(* IEC 61131-3 sources: 89152_FlorisHendrix_AfstudeerProject/89152_FlorisHendrix_ExamenProject/Stations/MachineControl/MachineControl/Network/HW_Network, 1 file *)

(* ---- ONE_HW_Network_Table.st ---- *)
#define OBJECTS_CONFIG

//Define part of class SdiasBase
//Address to access the Dataobject list via SPI SDO Read
#define SDIAS_SPI_DATA_OBJECT_LIST_PAGE_ADDRESS               16#FFFF
#define SDIAS_SPI_DATA_OBJECT_LIST_PAGE_OFFSET                16#00
#define SDIAS_SPI_DATA_OBJECT_LIST_IDENTIFIER                 16#12345678

//Defines the number of optional list elements in the SPI List

#define SDIAS_SPI_NUMBER_OF_OPTIONAL_ELEMENTS                 16

#define SDIAS_SPI_HEADER_BEFORE_OPTIONAL_ELEMENTS             16#18
#define SDIAS_SPI_HARDWARE_VERSION_OFFSET                     16#C
#define SDIAS_SPI_VENDOR_ID_OFFSET                            16#0

#define SDIAS_SPI_MASTER_ADRESS_TRANSMIT_BUFFER0              16#0000
#define SDIAS_SPI_MASTER_ADRESS_TRANSMIT_BUFFER1              16#0080
#define SDIAS_SPI_MASTER_ADRESS_RECEIVE_BUFFER0               16#0000
#define SDIAS_SPI_MASTER_ADRESS_RECEIVE_BUFFER1               16#0080
#define SDIAS_SPI_MASTER_ADRESS_PAGE_ADRESS                   16#0100
#define SDIAS_SPI_MASTER_ADRESS_PREDEFINED_COMMAND_REGISTER   16#0102
#define SDIAS_SPI_MASTER_ADRESS_SINGLE_COMMAND_REGISTER       16#0103
#define SDIAS_SPI_MASTER_ADRESS_STATUS_REGISTER               16#0104
#define SDIAS_SPI_MASTER_ADRESS_REQUEST_REGISTER              16#0105
#define SDIAS_SPI_MASTER_ADRESS_GRANT_REGISTER                16#0106
#define SDIAS_SPI_MASTER_ADRESS_CLEAR_REQUEST_REGISTER        16#0107
#define SDIAS_SPI_MASTER_ADRESS_FEATURE_REGISTER              16#0108

#define SDIAS_SPI_MASTER_SOFTWARE_REQUEST                     1

#define SDIAS_SPI_MASTER_COMMAND_PAGE_READ                    16#01
#define SDIAS_SPI_MASTER_COMMAND_PAGE_PROGRAM                 16#02
#define SDIAS_SPI_MASTER_COMMAND_SECTOR_ERASE                 16#03
#define SDIAS_SPI_MASTER_COMMAND_REBOOT_FPGA                  16#F0

#define SDIAS_SPI_MASTER_STATE_BUSY                           16#00
#define SDIAS_SPI_MASTER_STATE_READY                          16#01

#define SDIAS_SPI_SECTOR_SIZE                                 65536 // 256*256
#define SDIAS_SPI_PAGE_SIZE                                   256

#define SDIAS_SPI_WRITE_MAX_RETRIES                           2
#define SDIAS_SPI_TIMEOUT                                     500  //timeout for spi accesses
#define SDIAS_SPI_LOCK_TIMEOUT                                6   //this value is multiplied with the buscycletime [µs] (6*1000=6.000 msec timeout)

//SPI List IDs
#define SDIAS_SPI_IDENTIFICATION_LIST_ID  1
#define SDIAS_SPI_FLASH_CONFIGURATION_ID  2
#define SDIAS_SPI_VENDOR_NAME_ID          3
#define SDIAS_SPI_DEVICE_NAME_ID          4
#define SDIAS_SPI_SERIAL_NUMBER_ID        5
#define SDIAS_SPI_ORDERING_NUMBER_ID      6
#define SDIAS_SPI_DOCUMENTATION_PDF_ID    7
#define SDIAS_SPI_CALIB_DATA_ID           10
#define SDIAS_SPI_PDO_INFORMATION_ID      128

//SPI Access
#define SDIAS_SPI_ACCESS_ID_HW_TREE          1
#define SDIAS_SPI_ACCESS_ID_HWK_INTERNAL     2
#include "..\..\Class\SdiasManager\SdiasManager.h"
#include "..\..\Class\SdiasBase\SdiasBase.h"
#include "..\..\Class\HwControl\HwControl.h"
#include "..\..\Source\interfaces\lsl_st_hardwaretree.h"
#include "..\..\Source\interfaces\lsl_st_mt.h"
//Define part of class _BusInterfaceSdiasDriveMng
#define BUSIF_SDIASDRIVEMNG_OFFSET_TYPELABEL        0x0000
#define BUSIF_SDIASDRIVEMNG_PARALIST_INDEX_SET      0x2210
#define BUSIF_SDIASDRIVEMNG_PARALIST_INDEX_INFO     0x2211
#define BUSIF_SDIASDRIVEMNG_PARALIST_INDEX_SETNR    174

#define BUSIF_SDIASDRIVEMNG_MAX_SERVICEBOX          4
#define BUSIF_SDIASDRIVEMNG_SDO_RESPONSE_TIMEOUT    SDIAS_SDO_TIMEOUT * 2
#define BUSIF_SDIASDRIVEMNG_SDO_TYPELABEL_TIMEOUT   10000  //10 sec timeout to read typelabel

#define BUSIF_SDIASDRIVEMNG_SDO_SERVICE_APP_MDD100        0x4150
#define BUSIF_SDIASDRIVEMNG_SDO_SERVICE_APP_LASAL         0x4C41
#define BUSIF_SDIASDRIVEMNG_SDO_SERVICE_APP_CANOPEN       0x4453
#define BUSIF_SDIASDRIVEMNG_SDO_SERVICE_APP_CANOPEN_LASAL 0x444C

#define BUSIF_SDIASDRIVEMNG_FULL_PARADATA_SIZE   12
#define BUSIF_SDIASDRIVEMNG_CANOPEN_FOOTER_SIZE   4
#define BUSIF_SDIASDRIVEMNG_LASAL_PARADATA_SIZE   4

// if it's an sr011 or sr012 module we must set the pll system periode time with this offset
#define BUSIF_SDIASDRIVEMNG_SR01X_PLL_OFFSET    16#140
#include "..\..\class\_drivemngbase\drivemngbase.h"
//Define part of class _DriveAxisBase
// Device ID for the Drive Cards
#define DRIVEMNG_AXISDEVICEID_SDD_OFFSET         0
#define DRIVEMNG_AXISEVICEID_MDD_OFFSET   16#10000
#define DRIVEMNG_AXISEVICEID_SDIAS_OFFSET 16#20000

#define DRIVEAXIS_SPEED_SFFLIMITATION_USERINFO_0   32767
#define DRIVEAXIS_SPEED_SFFLIMITATION_USERINFO_1    1000
#define DRIVEAXIS_TORQUE_LIMITATION_VALUE           1000
#include "..\..\Class\_DriveMngBase\SDDDefinitions.h"
#include "..\..\Class\_DriveAxisBase\_DriveAxis_A_INT_Def.h"
//Define part of class _DriveMngBase
#ifndef _T_DRIVEMNGBASE_H
#define _T_DRIVEMNGBASE_H

// DiasDrive Constants
#DEFINE SDDMAXENTRIES   32        // maximale Anzahl an Achsen
#DEFINE SDDMAXPLACE     3         // maximale Anzahl an Achsen pro Steckplatz

// Device ID for the Drive IF Cards
#define DRIVEMNG_BUSDEVICEID_VAC011    11
#define DRIVEMNG_BUSDEVICEID_VAC012  1061
#define DRIVEMNG_BUSDEVICEID_VAC013  1075

#define DRIVEMNG_BUSDEVICEID_MDD     1071

// Device ID for the Drive Cards
#define DRIVEMNG_DRVDEVICEID_SDD_OFFSET 0

#define DRIVEMNG_DRVDEVICEID_SDD305 DRIVEMNG_DRVDEVICEID_SDD_OFFSET + 16
#define DRIVEMNG_DRVDEVICEID_SDD310 DRIVEMNG_DRVDEVICEID_SDD_OFFSET +  3
#define DRIVEMNG_DRVDEVICEID_SDD315 DRIVEMNG_DRVDEVICEID_SDD_OFFSET +  1
#define DRIVEMNG_DRVDEVICEID_SDD335 DRIVEMNG_DRVDEVICEID_SDD_OFFSET + 12

#define DRIVEMNG_DRVDEVICEID_SDD205 DRIVEMNG_DRVDEVICEID_SDD_OFFSET + 22
#define DRIVEMNG_DRVDEVICEID_SDD210 DRIVEMNG_DRVDEVICEID_SDD_OFFSET +  9
#define DRIVEMNG_DRVDEVICEID_SDD215 DRIVEMNG_DRVDEVICEID_SDD_OFFSET +  5

#define DRIVEMNG_DRVDEVICEID_SDD105 DRIVEMNG_DRVDEVICEID_SDD_OFFSET + 21
#define DRIVEMNG_DRVDEVICEID_SDD115 DRIVEMNG_DRVDEVICEID_SDD_OFFSET + 10
#define DRIVEMNG_DRVDEVICEID_SDD120 DRIVEMNG_DRVDEVICEID_SDD_OFFSET +  7

#define DRIVEMNG_DRVDEVICEID_MDD_OFFSET 16#10000

#define DRIVEMNG_DRVDEVICEID_MDD111 DRIVEMNG_DRVDEVICEID_MDD_OFFSET + 1
#define DRIVEMNG_DRVDEVICEID_MDD121 DRIVEMNG_DRVDEVICEID_MDD_OFFSET + 2

#define DRIVEMNG_DRVDEVICEID_SDIAS_OFFSET 16#20000

#define DRIVEMNG_DRVDEVICEID_DC061 DRIVEMNG_DRVDEVICEID_SDIAS_OFFSET + 16#180 // 1 = 1 Achse 80 SDIAS

#define DRIVEMNG_DRIVESCOPE_GETALL_PARAM    16#2080
#define DRIVEMNG_DRIVESCOPE_SCOPE_BIT       16#60000000
#define DRIVEMNG_DRIVESCOPE_SINDEX_RANGE    511

#define DRIVEMNG_DEFAULT_CPU_LOGFILENAME_PATH           "C:\sysmsg\DriveLog"
#define DRIVEMNG_DEFAULT_CPU_DEBUGLOGFILENAME_PATH      "C:\sysmsg\DriveDebugLog"
#define DRIVEMNG_DEFAULT_CPU_LOGFILENAME_EXTENSION      ".txt"

#define DRIVEMNG_DEFAULT_DRIVE_LOGFILENAME_PATH         "C:\"
#define DRIVEMNG_DEFAULT_DRIVE_LOGFILENAME_NAME         "DriveLog.txt"
#define DRIVEMNG_DEFAULT_DRIVE_DEBUGLOGFILENAME_NAME    "DriveDebugLog.txt"

#define DRIVEMNG_FILE_HANDLING_RETCODE_NOERROR                    0
#define DRIVEMNG_FILE_HANDLING_RETCODE_FILEHANDLING_BUSY         -2   // = DRIVEVVBASE_VANDAL_FILEHANDLING_ERROR_BUSY -2
#define DRIVEMNG_FILE_HANDLING_RETCODE_CMDVERSION_NOTSUPPORTED  -92
#define DRIVEMNG_FILE_HANDLING_RETCODE_WRITEPARA_FAILED         -93
#define DRIVEMNG_FILE_HANDLING_RETCODE_WRITEPARA_TIMEOUT        -94
#define DRIVEMNG_FILE_HANDLING_RETCODE_READBACKPARA_FAILED      -95
#define DRIVEMNG_FILE_HANDLING_RETCODE_READBACKPARA_TIMEOUT     -96
#define DRIVEMNG_FILE_HANDLING_RETCODE_AXIS_ENABLED             -97
#define DRIVEMNG_FILE_HANDLING_RETCODE_NOT_ONLINE               -98
#define DRIVEMNG_FILE_HANDLING_RETCODE_NOT_SUPPORTED            -99

#define DRIVEMNG_FILE_HANDLING_TIMEOUT_LOG_PARAM          10000

#define DRIVEMNG_FILESELECT_LOGFILE       0
#define DRIVEMNG_FILESELECT_DEBUGLOGFILE  1

#define DRIVEMNG_FILE_RESERVE_IDFREE         0
#define DRIVEMNG_FILE_RESERVE_IDDEFAULT     10
#define DRIVEMNG_FILE_RESERVE_IDGETLOGFILE  20

#endif // _T_DRIVEMNGBASE_H
//Define part of class AI043
#define DEVICE_ID_AI043 1045

#define AI043_ADDR_CYC_WRITE        16#000
#define AI043_ADDR_CYC_READ         16#080
#define AI043_ADDR_CFG_FIRMWARE     16#100
#define AI043_ADDR_STATE_FIRMWARE   16#180

#define AI043_SDO_RESPONSE_TIMEOUT  SDIAS_SDO_TIMEOUT * 2

#define AI043_KTY84_RAW_VALUES_FW_VER_AVAILABLE  16#110
#define AI043_AMOUNT_OF_VALID_CFG   25
#define AI043_AMOUNT_OF_VALID_CFGS_BEFORE_KTY84_ADDED 23

#define AI043_NUMBER_OF_ANALOG_IN   4
#define AI043_INVALID_VALUE         16#80000010$DINT
#define AI043_CABLE_BREAK_MASK      16#0F  //4 BITS

#define AI043_FIRMWARE_MIN          0
#define AI043_FIRMWARE_MAX_CFG12    2500
#define AI043_FIRMWARE_MAX_CFG13    5000
#define AI043_FIRMWARE_MAX_CFG14    10000
#define AI043_FIRMWARE_MAX_CFG15    25000
#define AI043_FIRMWARE_MAX_CFG16    50000
//Define part of class BusInterfaceSDIASInternal
#define BUSIF_INTERNAL_MAX_NR_DO 100

// Defines for Mutex Generation
#define INTERNAL_STR_MUTEX_NAME_SEPERATOR ".."
#define INTERNAL_MUTEX_NAME_END_LENGTH 5
#define INTERNAL_MUTEX_NAME_MAX_LENGTH 32
#include "..\..\Source\BusInterface.h"
//Define part of class Varan_Base
#ifndef _T_VARANBASE_H
#define _T_VARANBASE_H

#define	VARAN_PLL_OFFSET		16#0140
#define VARAN_MULTIPLE_OFFSET	16#01AC

// version of serial number validation (16#10 = 1.0)
#define SERNO_VALIDATION_VERSION 16#10

#define IsTransparent_IS_AVAILABLE

// Defines for Mutex Generation
#define VARAN_STR_MUTEX_NAME_SEPERATOR ".."
#define VARAN_MUTEX_NAME_END_LENGTH 5
#define VARAN_MUTEX_NAME_MAX_LENGTH 32

#define VARAN_SPI_IDENT_LICENCENO_OFFSET    16#14
#define VARAN_SPI_IDENT_HARDWAREVER_OFFSET  16#18

#endif // _T_VARANBASE_H
//Define part of class BusInterfaceVARAN
#define BUSIF_VARAN_MAX_NR_DO     100
#define BUSIF_VARAN_MAX_NR_MOVEDO 100

#define BUSIF_VARAN_MAX_SDO 1

#define BUSIF_VARAN_BUS_READY_VER 16#1109
#include "..\..\Source\interfaces\lsl_st_pci.h"
//Define part of class DM081
#define DEVICE_ID_DM081 1028
//Define part of class DM161
#define DEVICE_ID_DM161 1029
#include "..\..\Class\HwControl\watchdog.h"
#include "..\..\Source\interfaces\lsl_st_sysinfo.h"
#include "..\..\Source\interfaces\lsl_st_systrace.h"
#include "..\..\Class\HwControl\_HWKScope.h"
#include <.\lsl_st_mt.h>
//Define part of class SafetyUDP
#define SAFETY_UDP_MAX_SOCKETS                6     // Max number of socket

#define SAFETY_UDP_CLT_SEND_OK                0    // Send ok
#define SAFETY_UDP_CLT_INVALID_HANDLE        -1    // Invalid handle
#define SAFETY_UDP_CLT_NOT_OPEN              -2    // Socket is not open
#define SAFETY_UDP_CLT_SEND_FAILED           -3    // Send failed
#define SAFETY_UDP_CLT_SEND_BUFFER_FULL      -4    // Send buffer is full
#define SAFETY_UDP_CLT_DATA_TO_BIG           -5    // Data to big

#define SAFETY_UDP_MAXIMUM_SEGMENT_SIZE    1452    // Maximum of user data

#define SAFETY_UDP_TIMEOUT_OPENSOCKET    (1000)    //timeout for opening socket

#define SAFETY_UDP_RECEIVE_TIMEOUT          800

#define SAFETY_UDP_TX_BUFFER_SIZE          1024
//Define part of class SafetyManager
#define LogBufferSize 1000
#include "..\..\Class\SafetyManager\SafetyManager.h"
#include "..\..\Source\interfaces\lsl_st_safetydll.h"
//Define part of class SdiasManager
#define SDIAS_SDO_MAX_LENGTH              128
#define SDIAS_SDO_RINGBUFFER_NO            64
#define SDIAS_SDO_CHANNEL_NO                3   // fixed in the VI hardware to be 3

// watchdog trigger interval (after 130ms of no trigger the SDIAS HW goes into reset again and takes at least another 10ms to be ready again)
#define SDIAS_WATCHDOG_TRIGGER_TIME        40

// time needed by sdias modules to start up after the watchdog is triggered the first time in ms
#define SDIAS_HARDWARE_STARTUP_TIME        15

// sdias manager needs 2 ticks to handle event for read task (measure sync time)
#define SDIAS_SYNC_MEASURE_TICKS            2

// after activating the PLL SyncOut it takes 3 cycles until the SDIAS sync can be injected
#define SDIAS_CYCLES_WAIT_AFTER_SYNC_ENABLE 3

// wait 1 bus cycle at start to get valid numbers in the task info
#define SDIAS_TASKINFO_READY_TICKS          1

// time to wait (in ms) until other tasks in the same or lower priority than post init have done their stuff
#define SDIAS_WAIT_TIME_IN_POST_INIT        1

#define SIZE_PER_SDIAS_CLIENT               16#0400

// for far memory accesses: 1 module can hold maximum 256 1K blocks (0-255)
#define SDIAS_1K_BLOCK_NO                       256

// far memory accesses maximum length in bytes
#define SDIAS_MAX_SIZE_FAR_MEM_ACCESS           127

#define SDIAS_OFFSET_HW_CONFIG              16#FF00
#define SDIAS_OFFSET_TASK_EVENT_IDS         16#FF10
#define SDIAS_OFFSET_FEATURE_INFO           16#FF18
#define SDIAS_OFFSET_APPLI_LED_STATES       16#FF20
#define SDIAS_OFFSET_SYNC_INJECTION_CFG     16#FF3D
#define SDIAS_OFFSET_TRIGGER_UNIT_SETUP_0   16#FF41
#define SDIAS_OFFSET_TRIGGER_UNIT_SETUP_1   16#FF45
#define SDIAS_OFFSET_TASK_START_CFG_0       16#FF60
#define SDIAS_OFFSET_TASK_CONFIG_0          16#FF86
#define SDIAS_OFFSET_TASK_CONFIG_1          16#FF96
#define SDIAS_OFFSET_TASK_INFO_1            16#FF94
#define SDIAS_OFFSET_TASK_HANDSHAKE_1       16#FF9B
#define SDIAS_OFFSET_TASK_DURATION_TIME_1   16#FF9C
#define SDIAS_OFFSET_TASK_DURATION_TIME_2   16#FFAC
#define SDIAS_OFFSET_TASK_CONFIG_2          16#FFA6

#define SDIAS_RETRIES_ALLOWED         2

// mask to get global error flag out of message counter byte of SDO responses
#define SDIAS_MASK_GLOBAL_ERROR_FLAG        16#80

// mask to get message counter out of message counter byte of SDO responses
#define SDIAS_MASK_MESSAGE_COUNTER          16#3F

#define SDIAS_EVENT_MASK_ID_SYNC_OUT0       16#10
#define SDIAS_EVENT_MASK_ID_SYNC_OUT1       16#11
#define SDIAS_EVENT_MASK_ID_SYNC_OUT2       16#12
#define SDIAS_EVENT_MASK_ID_SYNC_OUT3       16#13

#define SDIAS_MANAGER_SYNC_SYNCOUT_ID       16#85
#define SDIAS_TASK_START_EVENT_SYNCOUT_ID   16#86

#define SDIAS_PLACE_NO_MODULE_ADDED_SO_FAR  16#80000000

#define SDIAS_TRIGGER_UNIT_BYTE_SIZE        2

#define SDIAS_WAIT_TIME_FIRMWARE_HANDSHAKE  5 * 1000

// if the firmware version is below this, there might be problems with SCP111 and other modules => print warning at startup
#define SDIAS_FW_VERSION_SDO_ERROR_FIXED    16#120

// if the protocol version ist below this, Control Read/Broadcast Write Command is not supported by sdiasmanager
#define SDIAS_PROTOCOLVERSION_BROADCAST     16#120

// if the cil version ist below this, Control Read/Broadcast Write Command is not supported by OS for local SDIAS.
#define SDIAS_CILVERSION_BROADCAST         16#5001

// timeout for blocking the init during initialisation (in ms)
#define SDIAS_INIT_BLOCK_TIMEOUT            20 * 1000

#define SDIAS_MUTEX_NAME_END_LENGTH 3
#define SDIAS_MUTEX_NAME_MAX_LENGTH 32
#define SDIAS_MUTEX_STR_SEPERATOR   ".."

//#define SDIAS_RT_TIME_MEASUREMENT
#ifdef SDIAS_RT_TIME_MEASUREMENT
  #pragma message("ATTENTION: SDIAS real time measurement is active and needs additional ressources in the realtime task")
#endif

(* SDIAS data object commands  *)
#define	 SDIAS_CMD_END							  0x00			(* End command										          *)
#define	 SDIAS_CMD_ACC_MEMORY				  0x01			(* Access dpram memory								      *)
#define	 SDIAS_CMD_ACC_CONTROL				0x02			(* Access dpram control memory						  *)
#define	 SDIAS_CMD_GLOBAL						  0x03			(* SDIAS global command								      *)
#define	 SDIAS_CMD_COPY_LOCAL					0x04			(* DPRAM copy command in local dpram				*)
#define	 SDIAS_CMD_JMP_LOCAL					0x05			(* DPRAM jump command in local dpram 				*)
#define  SDIAS_CMD_ACC_MEMORY_FAR     0x07      (* SDIAS Far Memory Access                  *)

(* SDIAS defines for data object handling *)
// Write data oject list
#define	 SDIAS_DOL_WRITE_USAGE_DOL_EMPTY	  0x20			(* Usage of empty write dol list (wachtdog trigger + end command)   *)
#define	 SDIAS_DOL_WRITE_USAGE_DTA_EMPTY	  0x03			(* Usage of empty write dol data (DO ctrl of 2x copy command for task information + DO ctrl of watchdog trigger      *)
#define	 SDIAS_DOL_WRITE_OFFSET_END_CMD			0x10			(* One data object in list - offset = 1 DO size = 0x10						  *)
#define	 SDIAS_DOL_WRITE_OFFSET_FIRST_DTA		0x02			(* Offset of first data byte of second copy command = 2 (DO ctrl)   *)
#define	 SDIAS_DOL_WRITE_OFFSET_LAST_DTA		0x02			(* Offset of last data byte of second copy command = 2 (DO ctrl )   *)

// Read data oject list
#define	 SDIAS_DOL_READ_USAGE_DOL_EMPTY	    0x30			(* Usage of empty read dol list (2x task info copy command + end command)   *)
#define	 SDIAS_DOL_READ_USAGE_DTA_EMPTY	    0x0D			(* Usage of empty write dol data (DO ctrl of 2x copy command for task information + DO ctrl of watchdog trigger      *)
#define	 SDIAS_DOL_READ_OFFSET_END_CMD			0x20			(* One data object in list - offset = 1 DO size = 0x10						          *)
#define	 SDIAS_DOL_READ_OFFSET_FIRST_DTA		0x07			(* Offset of first data byte of second copy command = 7 = DO state          *)
#define	 SDIAS_DOL_READ_OFFSET_LAST_DTA		  0x0C			(* Offset of last data byte of second copy command = 12 (last byte of task information)       *)

//Versionsnumber where SDIAS SPI Read Accesses are available
#define  SDIAS_SDO_SPI_FIRMWARE_VERSION_AVAILABLE 16#0120

//error info mask
#define  SDIAS_ERROR_INFO_MASK    2#1000011000011111

// Broadcast DO Info
#define SDIAS_OFFSET_CLIENT_CTRLTIMESTAMP   16#0190
#define SDIAS_NR_TIMEBROADCAST_DOS 2
#define SDIAS_TIMEBROADCAST_SUBCMD 16#B0
#include "..\..\source\interfaces\lsl_st_pll.h"
//Define part of class SdiasPLC
#define SDIASM_OBJECT_PATH            16#88000002   // Object Path for VSDIASmanager Length = 2 (First 2byte), Domain = 0 (3rd byte), Escape Sequence SDIAS (4th byte)
//Define part of class VaranManager
#define SIZE_PAYLOAD_FRAME_HEADER_DO      16#38  // Const because datasize is in the Payload DOs
#define SIZE_PAYLOAD_IRQ_FRAME_HEADER_DO  16#40  // Const because datasize is in the Payload DOs

#define VM_MAX_POST_INIT_MODULES  1000

#define VM_OBJECT_PATH            16#81000002   // Object Path for Varanmanager Length = 2 (First 2byte), Domain = 0 (3rd byte), Escape Sequence Varan (4th byte)
#include "..\..\Class\VaranManager\VaranManager.h"
#include "..\..\Source\interfaces\lsl_st_kernel.h"
//Define part of class VI021
#define DEVICE_ID_VI022 1233

FUNCTION GLOBAL TAB ONE_HW_Network
-1$UINT, 0$UINT,
0$UINT, 0$UINT,

40$UDINT,
TO_UDINT(1048633017), "_BusInterfaceSdiasDriveMng", 1$UINT, 14$UINT, 2$UINT,
TO_UDINT(529317953), "_CanLib", 1$UINT, 10$UINT, 2$UINT,
TO_UDINT(912370472), "_DriveAxis", 1$UINT, 72$UINT, 1$UINT,
TO_UDINT(4124502522), "_DriveAxisBase", 1$UINT, 81$UINT, 0$UINT,
TO_UDINT(833307860), "_DriveAxisSet", 1$UINT, 22$UINT, 1$UINT,
TO_UDINT(1470062879), "_DriveMng_DC062", 1$UINT, 82$UINT, 2$UINT,
TO_UDINT(496739206), "_DriveMngBase", 1$UINT, 61$UINT, 0$UINT,
TO_UDINT(4078275645), "_SerLib", 1$UINT, 34$UINT, 3$UINT,
TO_UDINT(1698489890), "AI043", 1$UINT, 20$UINT, 1$UINT,
TO_UDINT(2897291062), "ASCII_BIN", 1$UINT, 21$UINT, 1$UINT,
TO_UDINT(3882880897), "BusInterfaceSDIASInternal", 2$UINT, 1$UINT, 0$UINT,
TO_UDINT(24783181), "BusInterfaceVARAN", 1$UINT, 75$UINT, 0$UINT,
TO_UDINT(658879389), "CP112_IOs", 1$UINT, 1$UINT, 1$UINT,
TO_UDINT(794617671), "CriticalSection", 0$UINT, 4$UINT, 2$UINT,
TO_UDINT(1610993701), "DM081", 1$UINT, 13$UINT, 1$UINT,
TO_UDINT(4282685340), "DM161", 1$UINT, 14$UINT, 1$UINT,
TO_UDINT(3238133653), "Hub_Base", 1$UINT, 21$UINT, 1$UINT,
TO_UDINT(1770276445), "Hub_Base_Root", 2$UINT, 11$UINT, 1$UINT,
TO_UDINT(3078259981), "HwcLogging", 1$UINT, 0$UINT, 1$UINT,
TO_UDINT(2471641665), "HwControl", 5$UINT, 21$UINT, 1$UINT,
TO_UDINT(1193052171), "HwControlBase", 1$UINT, 10$UINT, 0$UINT,
TO_UDINT(4260294091), "HWRtPostScan", 1$UINT, 0$UINT, 1$UINT,
TO_UDINT(2225119864), "MerkerEx", 1$UINT, 22$UINT, 11$UINT,
TO_UDINT(933570811), "RAMex", 1$UINT, 17$UINT, 1$UINT,
TO_UDINT(3591333481), "RamFile", 1$UINT, 9$UINT, 1$UINT,
TO_UDINT(1799751072), "SafetyManager", 2$UINT, 26$UINT, 1$UINT,
TO_UDINT(3727715967), "SafetyUDP", 1$UINT, 4$UINT, 0$UINT,
TO_UDINT(3175101883), "SdiasBase", 1$UINT, 60$UINT, 0$UINT,
TO_UDINT(4173303375), "SdiasHubBase", 1$UINT, 10$UINT, 2$UINT,
TO_UDINT(2118381352), "SdiasManager", 1$UINT, 97$UINT, 2$UINT,
TO_UDINT(1159122596), "SdiasPLC", 2$UINT, 6$UINT, 1$UINT,
TO_UDINT(1850111279), "String", 1$UINT, 11$UINT, 10$UINT,
TO_UDINT(2898603620), "StringInternal", 1$UINT, 85$UINT, 0$UINT,
TO_UDINT(862125188), "Varan_Base", 2$UINT, 20$UINT, 0$UINT,
TO_UDINT(2940693151), "VaranManager", 3$UINT, 7$UINT, 0$UINT,
TO_UDINT(1989862026), "VaranManager_1", 2$UINT, 7$UINT, 1$UINT,
TO_UDINT(4035182347), "VaranManager_Base", 1$UINT, 26$UINT, 0$UINT,
TO_UDINT(262695706), "VI021", 1$UINT, 101$UINT, 1$UINT,
TO_UDINT(3232495061), "VirtualBaseInit", 1$UINT, 3$UINT, 0$UINT,
TO_UDINT(819479645), "XXXBase_IOs", 1$UINT, 1$UINT, 0$UINT,

1$UINT, TO_UDINT(1755887647), "_DRIVEMNG_DC0621\BUSINTERFACESDIASDRIVEMNG",
1$UINT, TO_UDINT(3678180828), "_DRIVEMNG_DC0622\BUSINTERFACESDIASDRIVEMNG",

1$UINT, TO_UDINT(3194356815), "CP112_IOS1\_BASE\_CANLIB1",
1$UINT, TO_UDINT(661607925), "CP112_IOS1\_BASE\_CANLIB2",

_NO_ATTR, TO_UDINT(794195804), "_DRIVEAXIS2",

1$UINT, TO_UDINT(1732231006), "_DRIVEAXIS2\SDDAXSET1",

_NO_ATTR, TO_UDINT(243498275), "_DRIVEMNG_DC0621",
_NO_ATTR, TO_UDINT(2542415001), "_DRIVEMNG_DC0622",

1$UINT, TO_UDINT(3879313428), "CP112_IOS1\_BASE\_SERLIB1",
1$UINT, TO_UDINT(2117136814), "CP112_IOS1\_BASE\_SERLIB2",
1$UINT, TO_UDINT(154648888), "CP112_IOS1\_BASE\_SERLIB3",

_NO_ATTR, TO_UDINT(1457099445), "AI0431",

1$UINT, TO_UDINT(3603645853), "VARANMANAGER_11\_BASE\ASCII_BIN1",

_NO_ATTR, TO_UDINT(222643709), "CP112_IOS1",

1$UINT, TO_UDINT(2972590922), "HWCONTROL1\SAFETYMANAGER\UDPRECEIVEDATA",
1$UINT, TO_UDINT(1868223583), "HWCONTROL1\SAFETYMANAGER\UDPSENDDATA",

_NO_ATTR, TO_UDINT(3367517728), "DM0811",

_NO_ATTR, TO_UDINT(2056942671), "DM1611",

1$UINT, TO_UDINT(658018123), "VI0211\HUB_BASE1",

1$UINT, TO_UDINT(1776428101), "VARANMANAGER_11\HUB_BASE_ROOT0",

1$UINT, TO_UDINT(3105254819), "HWCONTROL1\HWCLOGGING",

_NO_ATTR, TO_UDINT(2190789875), "HWCONTROL1",

1$UINT, TO_UDINT(1673205898), "HWCONTROL1\HWRTPOSTSCAN",

1$UINT, TO_UDINT(3111676623), "AI0431\_BASE\SERIALNOSTR\MERKEREX0",
1$UINT, TO_UDINT(3763871537), "DM0811\_BASE\SERIALNOSTR\MERKEREX0",
1$UINT, TO_UDINT(1089285877), "DM1611\_BASE\SERIALNOSTR\MERKEREX0",
1$UINT, TO_UDINT(1965133148), "VI0211\_BASE\_BASE\SERIALNOSTR\MERKEREX0",
1$UINT, TO_UDINT(2138211921), "_DRIVEAXIS2\MERKEREX2",
1$UINT, TO_UDINT(1361534785), "_DRIVEMNG_DC0621\BUSINTERFACESDIASDRIVEMNG\_BASE\SERIALNOSTR\MERKEREX0",
1$UINT, TO_UDINT(570430050), "_DRIVEMNG_DC0621\FWDATESTRING\MERKEREX0",
1$UINT, TO_UDINT(1339808896), "_DRIVEMNG_DC0621\FWNUMSTRING\MERKEREX0",
1$UINT, TO_UDINT(925076081), "_DRIVEMNG_DC0622\BUSINTERFACESDIASDRIVEMNG\_BASE\SERIALNOSTR\MERKEREX0",
1$UINT, TO_UDINT(2048834378), "_DRIVEMNG_DC0622\FWDATESTRING\MERKEREX0",
1$UINT, TO_UDINT(960423357), "_DRIVEMNG_DC0622\FWNUMSTRING\MERKEREX0",

1$UINT, TO_UDINT(1158084118), "_DRIVEAXIS2\RAMEX2",

1$UINT, TO_UDINT(4171808520), "VI0211\_BASE\_BASE\SERNOBACKUP",

1$UINT, TO_UDINT(1778590035), "HWCONTROL1\SAFETYMANAGER",

1$UINT, TO_UDINT(1007630054), "SDIASPLC1\SDIASHUBBASE1",
1$UINT, TO_UDINT(1199943557), "VI0211\SDIASHUBBASE",

1$UINT, TO_UDINT(4015996540), "SDIASPLC1\SDIASMANAGER1",
1$UINT, TO_UDINT(3245985506), "VI0211\SDIASMANAGER",

_NO_ATTR, TO_UDINT(1378000520), "SDIASPLC1",

1$UINT, TO_UDINT(2796855937), "AI0431\_BASE\SERIALNOSTR",
1$UINT, TO_UDINT(3004072747), "DM0811\_BASE\SERIALNOSTR",
1$UINT, TO_UDINT(2011818843), "DM1611\_BASE\SERIALNOSTR",
1$UINT, TO_UDINT(3053332208), "VI0211\_BASE\_BASE\SERIALNOSTR",
1$UINT, TO_UDINT(189353776), "_DRIVEMNG_DC0621\BUSINTERFACESDIASDRIVEMNG\_BASE\SERIALNOSTR",
1$UINT, TO_UDINT(275191107), "_DRIVEMNG_DC0621\FWDATESTRING",
1$UINT, TO_UDINT(1236665617), "_DRIVEMNG_DC0621\FWNUMSTRING",
1$UINT, TO_UDINT(880947621), "_DRIVEMNG_DC0622\BUSINTERFACESDIASDRIVEMNG\_BASE\SERIALNOSTR",
1$UINT, TO_UDINT(1812344984), "_DRIVEMNG_DC0622\FWDATESTRING",
1$UINT, TO_UDINT(4101794271), "_DRIVEMNG_DC0622\FWNUMSTRING",

_NO_ATTR, TO_UDINT(2395414379), "VARANMANAGER_11",

_NO_ATTR, TO_UDINT(2125577894), "VI0211",

//Internal connections
0$UDINT,
43$UDINT,
TO_UDINT(0), "SerialNoStr", TO_UDINT(46),
TO_UDINT(1), "SerialNoStr", TO_UDINT(49),
TO_UDINT(4), "SDDAxSet1", TO_UDINT(5),
TO_UDINT(4), "MerkerEx2", TO_UDINT(27),
TO_UDINT(4), "RAMex2", TO_UDINT(34),
TO_UDINT(6), "FWDateString", TO_UDINT(47),
TO_UDINT(6), "FWNumSTring", TO_UDINT(48),
TO_UDINT(6), "BusInterfaceSdiasDriveMng", TO_UDINT(0),
TO_UDINT(7), "FWDateString", TO_UDINT(50),
TO_UDINT(7), "FWNumSTring", TO_UDINT(51),
TO_UDINT(7), "BusInterfaceSdiasDriveMng", TO_UDINT(1),
TO_UDINT(11), "SerialNoStr", TO_UDINT(42),
TO_UDINT(13), "_SerLib1", TO_UDINT(8),
TO_UDINT(13), "_SerLib2", TO_UDINT(9),
TO_UDINT(13), "_CanLib1", TO_UDINT(2),
TO_UDINT(13), "_CanLib2", TO_UDINT(3),
TO_UDINT(13), "_SerLib3", TO_UDINT(10),
TO_UDINT(16), "SerialNoStr", TO_UDINT(43),
TO_UDINT(17), "SerialNoStr", TO_UDINT(44),
TO_UDINT(21), "SafetyManager", TO_UDINT(36),
TO_UDINT(21), "HWRtPostScan", TO_UDINT(22),
TO_UDINT(21), "HwcLogging", TO_UDINT(20),
TO_UDINT(36), "UdpSendData", TO_UDINT(15),
TO_UDINT(36), "UdpReceiveData", TO_UDINT(14),
TO_UDINT(41), "SdiasManager1", TO_UDINT(39),
TO_UDINT(41), "SdiasHubBase1", TO_UDINT(37),
TO_UDINT(42), "MerkerEx0", TO_UDINT(23),
TO_UDINT(43), "MerkerEx0", TO_UDINT(24),
TO_UDINT(44), "MerkerEx0", TO_UDINT(25),
TO_UDINT(45), "MerkerEx0", TO_UDINT(26),
TO_UDINT(46), "MerkerEx0", TO_UDINT(28),
TO_UDINT(47), "MerkerEx0", TO_UDINT(29),
TO_UDINT(48), "MerkerEx0", TO_UDINT(30),
TO_UDINT(49), "MerkerEx0", TO_UDINT(31),
TO_UDINT(50), "MerkerEx0", TO_UDINT(32),
TO_UDINT(51), "MerkerEx0", TO_UDINT(33),
TO_UDINT(52), "ASCII_BIN1", TO_UDINT(12),
TO_UDINT(52), "Hub_Base_Root0", TO_UDINT(19),
TO_UDINT(53), "SerialNoStr", TO_UDINT(45),
TO_UDINT(53), "SerNoBackup", TO_UDINT(35),
TO_UDINT(53), "Hub_Base1", TO_UDINT(18),
TO_UDINT(53), "SdiasManager", TO_UDINT(40),
TO_UDINT(53), "SdiasHubBase", TO_UDINT(38),
0$UDINT,
39$UDINT,
TO_UDINT(4), "DriveMng", TO_UDINT(7), "CmdState",
TO_UDINT(4), "DriveAxisSet", TO_UDINT(5), "Server0",
TO_UDINT(5), "coMerkerEx", TO_UDINT(27), "m_udLength",
TO_UDINT(5), "coRamEx", TO_UDINT(34), "m_udLength",
TO_UDINT(6), "cOnline", TO_UDINT(0), "Online",
TO_UDINT(6), "FwNumStr", TO_UDINT(48), "Data",
TO_UDINT(6), "FwDatetr", TO_UDINT(47), "Data",
TO_UDINT(6), "ToBusIF", TO_UDINT(0), "CallCommand",
TO_UDINT(6), "SdiasIn", TO_UDINT(38), "ClassSvr",
TO_UDINT(7), "cOnline", TO_UDINT(1), "Online",
TO_UDINT(7), "FwNumStr", TO_UDINT(51), "Data",
TO_UDINT(7), "FwDatetr", TO_UDINT(50), "Data",
TO_UDINT(7), "ToBusIF", TO_UDINT(1), "CallCommand",
TO_UDINT(7), "SdiasIn", TO_UDINT(38), "ClassSvr",
TO_UDINT(11), "SdiasIn", TO_UDINT(37), "ClassSvr",
TO_UDINT(13), "To_HwControl", TO_UDINT(21), "Control",
TO_UDINT(16), "SdiasIn", TO_UDINT(38), "ClassSvr",
TO_UDINT(17), "SdiasIn", TO_UDINT(37), "ClassSvr",
TO_UDINT(18), "VaranIn", TO_UDINT(53), "State",
TO_UDINT(19), "VaranConnect", TO_UDINT(52), "Control",
TO_UDINT(22), "toHwControlBase", TO_UDINT(21), "Control",
TO_UDINT(36), "To_HwControl", TO_UDINT(21), "Control",
TO_UDINT(37), "ToNextSDIAS", TO_UDINT(39), "ClassState",
TO_UDINT(38), "ToNextSDIAS", TO_UDINT(40), "ClassState",
TO_UDINT(39), "ToBusInterface", TO_UDINT(41), "CallCommand",
TO_UDINT(40), "ToBusInterface", TO_UDINT(53), "CallCommand",
TO_UDINT(41), "ToHwControl", TO_UDINT(21), "Control",
TO_UDINT(42), "DataBuffer", TO_UDINT(23), "m_udLength",
TO_UDINT(43), "DataBuffer", TO_UDINT(24), "m_udLength",
TO_UDINT(44), "DataBuffer", TO_UDINT(25), "m_udLength",
TO_UDINT(45), "DataBuffer", TO_UDINT(26), "m_udLength",
TO_UDINT(46), "DataBuffer", TO_UDINT(28), "m_udLength",
TO_UDINT(47), "DataBuffer", TO_UDINT(29), "m_udLength",
TO_UDINT(48), "DataBuffer", TO_UDINT(30), "m_udLength",
TO_UDINT(49), "DataBuffer", TO_UDINT(31), "m_udLength",
TO_UDINT(50), "DataBuffer", TO_UDINT(32), "m_udLength",
TO_UDINT(51), "DataBuffer", TO_UDINT(33), "m_udLength",
TO_UDINT(52), "To_HwControl", TO_UDINT(21), "Control",
TO_UDINT(53), "VaranIn", TO_UDINT(19), "Control",

//Initialization values
0$UDINT,
91$UDINT,
TO_UDINT(0), "LEDControl", TO_UDINT(0),//|HW_Network._DriveMng_DC0621\BusInterfaceSdiasDriveMng.LEDControl;
TO_UDINT(0), "Place", TO_UDINT(1),//|HW_Network._DriveMng_DC0621\BusInterfaceSdiasDriveMng.Place;
TO_UDINT(0), "Required", TO_UDINT(1),//|HW_Network._DriveMng_DC0621\BusInterfaceSdiasDriveMng.Required;
TO_UDINT(0), "TimeMultiplier", TO_UDINT(1),//|HW_Network._DriveMng_DC0621\BusInterfaceSdiasDriveMng.TimeMultiplier;
TO_UDINT(0), "SdiasID", TO_UDINT(1801),//|HW_Network._DriveMng_DC0621\BusInterfaceSdiasDriveMng.SdiasID;
TO_UDINT(1), "LEDControl", TO_UDINT(0),//|HW_Network._DriveMng_DC0622\BusInterfaceSdiasDriveMng.LEDControl;
TO_UDINT(1), "Place", TO_UDINT(2),//|HW_Network._DriveMng_DC0622\BusInterfaceSdiasDriveMng.Place;
TO_UDINT(1), "Required", TO_UDINT(1),//|HW_Network._DriveMng_DC0622\BusInterfaceSdiasDriveMng.Required;
TO_UDINT(1), "TimeMultiplier", TO_UDINT(1),//|HW_Network._DriveMng_DC0622\BusInterfaceSdiasDriveMng.TimeMultiplier;
TO_UDINT(1), "SdiasID", TO_UDINT(1801),//|HW_Network._DriveMng_DC0622\BusInterfaceSdiasDriveMng.SdiasID;
TO_UDINT(2), "CanBus", TO_UDINT(1),//|HW_Network._base\CP112_IOs1\_CanLib1.CanBus;
TO_UDINT(3), "CanBus", TO_UDINT(2),//|HW_Network._base\CP112_IOs1\_CanLib2.CanBus;
TO_UDINT(4), "Place", TO_UDINT(0),//|HW_Network._DriveAxis2.Place;
TO_UDINT(4), "AxisNo", TO_UDINT(1),//|HW_Network._DriveAxis2.AxisNo;
TO_UDINT(4), "AxisExtend", TO_UDINT(1),//|HW_Network._DriveAxis2.AxisExtend;
TO_UDINT(4), "ParaSaveType", TO_UDINT(1),//|HW_Network._DriveAxis2.ParaSaveType;
TO_UDINT(4), "OverwriteMotorPara", TO_UDINT(0),//|HW_Network._DriveAxis2.OverwriteMotorPara;
TO_UDINT(5), "ParaSaveType", TO_UDINT(1),//|HW_Network._DriveAxis2\SDDAxSet1.ParaSaveType;
TO_UDINT(5), "OverwriteMotorPara", TO_UDINT(0),//|HW_Network._DriveAxis2\SDDAxSet1.OverwriteMotorPara;
TO_UDINT(6), "Place", TO_UDINT(1),//|HW_Network._DriveMng_DC0621.Place;
TO_UDINT(6), "Required", TO_UDINT(1),//|HW_Network._DriveMng_DC0621.Required;
TO_UDINT(6), "TimeMultiplier", TO_UDINT(1),//|HW_Network._DriveMng_DC0621.TimeMultiplier;
TO_UDINT(7), "Place", TO_UDINT(2),//|HW_Network._DriveMng_DC0622.Place;
TO_UDINT(7), "Required", TO_UDINT(1),//|HW_Network._DriveMng_DC0622.Required;
TO_UDINT(7), "TimeMultiplier", TO_UDINT(1),//|HW_Network._DriveMng_DC0622.TimeMultiplier;
TO_UDINT(8), "Com", TO_UDINT(1),//|HW_Network._base\CP112_IOs1\_SerLib1.Com;
TO_UDINT(9), "Com", TO_UDINT(2),//|HW_Network._base\CP112_IOs1\_SerLib2.Com;
TO_UDINT(10), "Com", TO_UDINT(3),//|HW_Network._base\CP112_IOs1\_SerLib3.Com;
TO_UDINT(11), "LEDControl", TO_UDINT(0),//|HW_Network.AI0431.LEDControl;
TO_UDINT(11), "Place", TO_UDINT(1),//|HW_Network.AI0431.Place;
TO_UDINT(11), "Required", TO_UDINT(1),//|HW_Network.AI0431.Required;
TO_UDINT(11), "AI1_Active", TO_UDINT(1),//|HW_Network.AI0431.AI1_Active;
TO_UDINT(11), "AI2_Active", TO_UDINT(1),//|HW_Network.AI0431.AI2_Active;
TO_UDINT(11), "AI3_Active", TO_UDINT(1),//|HW_Network.AI0431.AI3_Active;
TO_UDINT(11), "AI4_Active", TO_UDINT(1),//|HW_Network.AI0431.AI4_Active;
TO_UDINT(16), "LEDControl", TO_UDINT(0),//|HW_Network.DM0811.LEDControl;
TO_UDINT(16), "Place", TO_UDINT(0),//|HW_Network.DM0811.Place;
TO_UDINT(16), "Required", TO_UDINT(1),//|HW_Network.DM0811.Required;
TO_UDINT(17), "LEDControl", TO_UDINT(0),//|HW_Network.DM1611.LEDControl;
TO_UDINT(17), "Place", TO_UDINT(0),//|HW_Network.DM1611.Place;
TO_UDINT(17), "Required", TO_UDINT(1),//|HW_Network.DM1611.Required;
TO_UDINT(18), "Splitter_Place", TO_UDINT(0),//|HW_Network.VI0211\Hub_Base1.Splitter_Place;
TO_UDINT(19), "Splitter_Place", TO_UDINT(0),//|HW_Network.VaranManager_11\Hub_Base_Root0.Splitter_Place;
TO_UDINT(21), "UdpSafetyPort", TO_UDINT(10823),//|HW_Network.HwControl1.UdpSafetyPort;
TO_UDINT(21), "InterfaceNo", TO_UDINT(1),//|HW_Network.HwControl1.InterfaceNo;
TO_UDINT(21), "RtTaskSync", TO_UDINT(0),//|HW_Network.HwControl1.RtTaskSync;
TO_UDINT(23), "ThreadSafe", TO_UDINT(0),//|HW_Network.SerialNoStr\_base\AI0431\MerkerEx0.ThreadSafe;
TO_UDINT(24), "ThreadSafe", TO_UDINT(0),//|HW_Network.SerialNoStr\_base\DM0811\MerkerEx0.ThreadSafe;
TO_UDINT(25), "ThreadSafe", TO_UDINT(0),//|HW_Network.SerialNoStr\_base\DM1611\MerkerEx0.ThreadSafe;
TO_UDINT(26), "ThreadSafe", TO_UDINT(0),//|HW_Network.SerialNoStr\_base\_base\VI0211\MerkerEx0.ThreadSafe;
TO_UDINT(27), "ThreadSafe", TO_UDINT(0),//|HW_Network._DriveAxis2\MerkerEx2.ThreadSafe;
TO_UDINT(28), "ThreadSafe", TO_UDINT(0),//|HW_Network.SerialNoStr\_base\BusInterfaceSdiasDriveMng\_DriveMng_DC0621\MerkerEx0.ThreadSafe;
TO_UDINT(29), "ThreadSafe", TO_UDINT(0),//|HW_Network.FWDateString\_DriveMng_DC0621\MerkerEx0.ThreadSafe;
TO_UDINT(30), "ThreadSafe", TO_UDINT(0),//|HW_Network.FWNumSTring\_DriveMng_DC0621\MerkerEx0.ThreadSafe;
TO_UDINT(31), "ThreadSafe", TO_UDINT(0),//|HW_Network.SerialNoStr\_base\BusInterfaceSdiasDriveMng\_DriveMng_DC0622\MerkerEx0.ThreadSafe;
TO_UDINT(32), "ThreadSafe", TO_UDINT(0),//|HW_Network.FWDateString\_DriveMng_DC0622\MerkerEx0.ThreadSafe;
TO_UDINT(33), "ThreadSafe", TO_UDINT(0),//|HW_Network.FWNumSTring\_DriveMng_DC0622\MerkerEx0.ThreadSafe;
TO_UDINT(34), "ThreadSafe", TO_UDINT(0),//|HW_Network._DriveAxis2\RAMex2.ThreadSafe;
TO_UDINT(35), "Setup", TO_UDINT(2#1101),//|HW_Network._base\_base\VI0211\SerNoBackup.Setup;
TO_UDINT(36), "UdpSafetyPort", TO_UDINT(10823),//|HW_Network.HwControl1\SafetyManager.UdpSafetyPort;
TO_UDINT(36), "InterfaceNo", TO_UDINT(1),//|HW_Network.HwControl1\SafetyManager.InterfaceNo;
TO_UDINT(36), "UdpSafetyRequestCycle", TO_UDINT(UDP_MIN_REQUEST_TIME),//|HW_Network.HwControl1\SafetyManager.UdpSafetyRequestCycle;
TO_UDINT(36), "UdpSafetyResponseTimeout", TO_UDINT(UDP_MIN_RESPONSE_TIMEOUT),//|HW_Network.HwControl1\SafetyManager.UdpSafetyResponseTimeout;
TO_UDINT(37), "SplitterPlace", TO_UDINT(0),//|HW_Network.SdiasPLC1\SdiasHubBase1.SplitterPlace;
TO_UDINT(38), "SplitterPlace", TO_UDINT(0),//|HW_Network.VI0211\SdiasHubBase.SplitterPlace;
TO_UDINT(39), "DeviceID", TO_UDINT(0),//|HW_Network.SdiasPLC1\SdiasManager1.DeviceID;
TO_UDINT(39), "AutoFarMem", TO_UDINT(0),//|HW_Network.SdiasPLC1\SdiasManager1.AutoFarMem;
TO_UDINT(40), "DeviceID", TO_UDINT(1187),//|HW_Network.VI0211\SdiasManager.DeviceID;
TO_UDINT(40), "AutoFarMem", TO_UDINT(0),//|HW_Network.VI0211\SdiasManager.AutoFarMem;
TO_UDINT(41), "CycleTime", TO_UDINT(1000),//|HW_Network.SdiasPLC1.CycleTime;
TO_UDINT(41), "IsoStartPoint", TO_UDINT(50),//|HW_Network.SdiasPLC1.IsoStartPoint;
TO_UDINT(41), "AutoFarMem", TO_UDINT(0),//|HW_Network.SdiasPLC1.AutoFarMem;
TO_UDINT(42), "SingleRealloc", TO_UDINT(1),//|HW_Network._base\AI0431\SerialNoStr.SingleRealloc;
TO_UDINT(43), "SingleRealloc", TO_UDINT(1),//|HW_Network._base\DM0811\SerialNoStr.SingleRealloc;
TO_UDINT(44), "SingleRealloc", TO_UDINT(1),//|HW_Network._base\DM1611\SerialNoStr.SingleRealloc;
TO_UDINT(45), "SingleRealloc", TO_UDINT(1),//|HW_Network._base\_base\VI0211\SerialNoStr.SingleRealloc;
TO_UDINT(46), "SingleRealloc", TO_UDINT(1),//|HW_Network._base\BusInterfaceSdiasDriveMng\_DriveMng_DC0621\SerialNoStr.SingleRealloc;
TO_UDINT(47), "SingleRealloc", TO_UDINT(1),//|HW_Network._DriveMng_DC0621\FWDateString.SingleRealloc;
TO_UDINT(48), "SingleRealloc", TO_UDINT(1),//|HW_Network._DriveMng_DC0621\FWNumSTring.SingleRealloc;
TO_UDINT(49), "SingleRealloc", TO_UDINT(1),//|HW_Network._base\BusInterfaceSdiasDriveMng\_DriveMng_DC0622\SerialNoStr.SingleRealloc;
TO_UDINT(50), "SingleRealloc", TO_UDINT(1),//|HW_Network._DriveMng_DC0622\FWDateString.SingleRealloc;
TO_UDINT(51), "SingleRealloc", TO_UDINT(1),//|HW_Network._DriveMng_DC0622\FWNumSTring.SingleRealloc;
TO_UDINT(52), "VaranManagerTime", TO_UDINT(1000000),//|HW_Network.VaranManager_11.VaranManagerTime;
TO_UDINT(52), "VaranManagerNr", TO_UDINT(0),//|HW_Network.VaranManager_11.VaranManagerNr;
TO_UDINT(52), "PayloadFrame", TO_UDINT(0),//|HW_Network.VaranManager_11.PayloadFrame;
TO_UDINT(52), "CoreSelect", TO_UDINT(0),//|HW_Network.VaranManager_11.CoreSelect;
TO_UDINT(52), "InterframeGap", TO_UDINT(0),//|HW_Network.VaranManager_11.InterframeGap;
TO_UDINT(53), "Required", TO_UDINT(1),//|HW_Network.VI0211.Required;
TO_UDINT(53), "Transparent", TO_UDINT(0),//|HW_Network.VI0211.Transparent;
TO_UDINT(53), "TimeBase", TO_UDINT(0),//|HW_Network.VI0211.TimeBase;
TO_UDINT(53), "TimeBaseOffset", TO_UDINT(0),//|HW_Network.VI0211.TimeBaseOffset;

//Symbolic initialization values
0$UDINT,
0$UDINT,

//Initialization of string values
0$UDINT,
0$UDINT,

//Configuration of tasks (RealTime, Cyclic, Background)
0$UDINT,
1$UDINT,
TO_UDINT(22), (1)$UDINT, 4194304$DINT, 	//HWCONTROL1\HWRTPOSTSCAN

0$UDINT,
2$UDINT,
TO_UDINT(6), (10)$UDINT, 4194303$DINT, 	//_DRIVEMNG_DC0621
TO_UDINT(7), (10)$UDINT, 4194303$DINT, 	//_DRIVEMNG_DC0622

0$UDINT,
0$UDINT,

//External connections
0$UDINT,
0$UDINT,

//Magic internal connections
0$UDINT,
17$UDINT,
TO_UDINT(0), "SdiasIn", TO_UDINT(6), "SdiasIn",
TO_UDINT(0), "Place", TO_UDINT(6), "Place",
TO_UDINT(0), "Required", TO_UDINT(6), "Required",
TO_UDINT(0), "TimeMultiplier", TO_UDINT(6), "TimeMultiplier",
TO_UDINT(1), "SdiasIn", TO_UDINT(7), "SdiasIn",
TO_UDINT(1), "Place", TO_UDINT(7), "Place",
TO_UDINT(1), "Required", TO_UDINT(7), "Required",
TO_UDINT(1), "TimeMultiplier", TO_UDINT(7), "TimeMultiplier",
TO_UDINT(5), "ParaSaveType", TO_UDINT(4), "ParaSaveType",
TO_UDINT(5), "OverwriteMotorPara", TO_UDINT(4), "OverwriteMotorPara",
TO_UDINT(5), "ParaTab", TO_UDINT(4), "ParaTab",
TO_UDINT(5), "FileHandle", TO_UDINT(4), "FileHandle",
TO_UDINT(5), "TableIndex", TO_UDINT(4), "TableIndex",
TO_UDINT(36), "UdpSafetyPort", TO_UDINT(21), "UdpSafetyPort",
TO_UDINT(36), "InterfaceNo", TO_UDINT(21), "InterfaceNo",
TO_UDINT(36), "SafetyDomainTimeout", TO_UDINT(21), "SafetyDomainTimeout",
TO_UDINT(39), "AutoFarMem", TO_UDINT(41), "AutoFarMem",

//Configuration of timeslots of tasks (RealTime, Cyclic)
#ifdef __LSLLDR_TIMESLOTS__
0$UDINT,
0$UDINT,

0$UDINT,
0$UDINT,

#endif //__LSLLDR_TIMESLOTS__

//MultiMaster connections
#ifdef __LSLLDR_MULTIMASTER__
0$UDINT,
0$UDINT,
#endif //__LSLLDR_MULTIMASTER__

//Configuration for task ID (RealTime, CyclicTime)
#ifdef __LSLLDR_TASKID__
"\\\\TASKS2  "
0$UDINT,
1$UDINT,
(0)$UDINT, 	//HWCONTROL1\HWRTPOSTSCAN

0$UDINT,
2$UDINT,
(0)$UDINT, 	//_DRIVEMNG_DC0621
(0)$UDINT, 	//_DRIVEMNG_DC0622

0$UDINT,
0$UDINT,

#endif //__LSLLDR_TASKID__

END_FUNCTION
